FUNCTION "PDH_J_Raw" : Void
{ S7_Optimized_Access := 'TRUE' }
VERSION : 0.1
//Erzeugt vom PDH (PDH-Test) am 2026-11-15 10:00 UTC – bei Änderungen im PDH neu herunterladen.
//Datenbaustein "Daten", Variante mit Siemens-Bibliothek LMQTT (TLS möglich), S7-1500, höchstens 1024 Byte je Nachricht.
//Schreibt feste Zeichen (UTF-8) ab buf[pos]. Passt es nicht, wird ovf gesetzt und nichts geschrieben.
   VAR_INPUT
      s : String;
   END_VAR

   VAR_IN_OUT
      buf : Array[*] of Byte;
      pos : DInt;
      ovf : Bool;
   END_VAR

   VAR_TEMP
      i : Int;
      n : Int;
   END_VAR


BEGIN
	IF #ovf THEN
	    RETURN;
	END_IF;
	#n := LEN(#s);
	IF #pos < LOWER_BOUND(ARR := #buf, DIM := 1) OR #pos + INT_TO_DINT(#n) - 1 > UPPER_BOUND(ARR := #buf, DIM := 1) THEN
	    #ovf := TRUE;
	    RETURN;
	END_IF;
	FOR #i := 1 TO #n DO
	    #buf[#pos] := CHAR_TO_BYTE(#s[#i]);
	    #pos := #pos + 1;
	END_FOR;
END_FUNCTION

FUNCTION "PDH_J_DInt" : Void
{ S7_Optimized_Access := 'TRUE' }
VERSION : 0.1
//Erzeugt vom PDH (PDH-Test) am 2026-11-15 10:00 UTC – bei Änderungen im PDH neu herunterladen.
//Datenbaustein "Daten", Variante mit Siemens-Bibliothek LMQTT (TLS möglich), S7-1500, höchstens 1024 Byte je Nachricht.
//Schreibt v als Dezimalzahl (auch -2147483648).
   VAR_INPUT
      v : DInt;
   END_VAR

   VAR_IN_OUT
      buf : Array[*] of Byte;
      pos : DInt;
      ovf : Bool;
   END_VAR

   VAR_TEMP
      x : DInt;
      d : DInt;
      k : Int;
      i : Int;
      need : DInt;
      dig : Array[0..9] of Byte;
   END_VAR


BEGIN
	IF #ovf THEN
	    RETURN;
	END_IF;
	// Ziffern rückwärts sammeln, ohne das Vorzeichen umzudrehen (sonst Überlauf bei -2147483648)
	#x := #v;
	#k := 0;
	REPEAT
	    #d := #x MOD 10;
	    IF #d < 0 THEN
	        #d := -#d;
	    END_IF;
	    #dig[#k] := DINT_TO_BYTE(#d + 48);
	    #k := #k + 1;
	    #x := #x / 10;
	UNTIL #x = 0
	END_REPEAT;
	#need := INT_TO_DINT(#k);
	IF #v < 0 THEN
	    #need := #need + 1;
	END_IF;
	IF #pos < LOWER_BOUND(ARR := #buf, DIM := 1) OR #pos + #need - 1 > UPPER_BOUND(ARR := #buf, DIM := 1) THEN
	    #ovf := TRUE;
	    RETURN;
	END_IF;
	IF #v < 0 THEN
	    #buf[#pos] := 16#2D;   // -
	    #pos := #pos + 1;
	END_IF;
	FOR #i := #k - 1 TO 0 BY -1 DO
	    #buf[#pos] := #dig[#i];
	    #pos := #pos + 1;
	END_FOR;
END_FUNCTION

FUNCTION "PDH_J_UDInt" : Void
{ S7_Optimized_Access := 'TRUE' }
VERSION : 0.1
//Erzeugt vom PDH (PDH-Test) am 2026-11-15 10:00 UTC – bei Änderungen im PDH neu herunterladen.
//Datenbaustein "Daten", Variante mit Siemens-Bibliothek LMQTT (TLS möglich), S7-1500, höchstens 1024 Byte je Nachricht.
//Schreibt v als Dezimalzahl ohne Vorzeichen.
   VAR_INPUT
      v : UDInt;
   END_VAR

   VAR_IN_OUT
      buf : Array[*] of Byte;
      pos : DInt;
      ovf : Bool;
   END_VAR

   VAR_TEMP
      x : UDInt;
      k : Int;
      i : Int;
      dig : Array[0..9] of Byte;
   END_VAR


BEGIN
	IF #ovf THEN
	    RETURN;
	END_IF;
	#x := #v;
	#k := 0;
	REPEAT
	    #dig[#k] := UDINT_TO_BYTE(#x MOD 10 + 48);
	    #k := #k + 1;
	    #x := #x / 10;
	UNTIL #x = 0
	END_REPEAT;
	IF #pos < LOWER_BOUND(ARR := #buf, DIM := 1) OR #pos + INT_TO_DINT(#k) - 1 > UPPER_BOUND(ARR := #buf, DIM := 1) THEN
	    #ovf := TRUE;
	    RETURN;
	END_IF;
	FOR #i := #k - 1 TO 0 BY -1 DO
	    #buf[#pos] := #dig[#i];
	    #pos := #pos + 1;
	END_FOR;
END_FUNCTION

FUNCTION "PDH_J_Num" : Void
{ S7_Optimized_Access := 'TRUE' }
VERSION : 0.1
//Erzeugt vom PDH (PDH-Test) am 2026-11-15 10:00 UTC – bei Änderungen im PDH neu herunterladen.
//Datenbaustein "Daten", Variante mit Siemens-Bibliothek LMQTT (TLS möglich), S7-1500, höchstens 1024 Byte je Nachricht.
//Schreibt x mit digits gültigen Stellen wie Go strconv.FormatFloat(x, 'E', digits - 1, …):
//[-]d.ddd…E±XX, Exponent mit mindestens zwei Ziffern. NaN, ±unendlich und Beträge über maxAbs als null.
//Gerundet wird zur nächsten Zahl, bei genau der Mitte zur geraden. Für Beträge von 1E-8 bis 1E36
//wird der Rundungsfehler exakt mitgerechnet (Dekker); außerhalb kann die letzte Stelle selten abweichen.
//Gleich halten mit sclNum in generate_test.go (Go-Nachbau dieses Ablaufs).
   VAR_INPUT
      x : LReal;
      digits : Int;   // 7 für Real, 15 für LReal
      maxAbs : LReal;   // größter Betrag, der als Zahl geschrieben wird
   END_VAR

   VAR_IN_OUT
      buf : Array[*] of Byte;
      pos : DInt;
      ovf : Bool;
   END_VAR

   VAR_TEMP
      a : LReal;
      t : LReal;
      s : LReal;
      p : LReal;
      y : LReal;
      lo : LReal;
      n : LReal;
      f : LReal;
      top : LReal;
      c : LReal;
      ah : LReal;
      al : LReal;
      bh : LReal;
      bl : LReal;
      ph : LReal;
      e : Int;
      k : Int;
      j : Int;
      i : Int;
      pass : Int;
      hiD : DInt;
      loD : DInt;
      neg : Bool;
      exact : Bool;
      odd : Bool;
      dig : Array[1..15] of Byte;
   END_VAR


BEGIN
	IF #ovf THEN
	    RETURN;
	END_IF;
	IF #digits < 1 OR #digits > 15 OR #pos < LOWER_BOUND(ARR := #buf, DIM := 1) OR #pos + INT_TO_DINT(#digits) + 6 > UPPER_BOUND(ARR := #buf, DIM := 1) THEN
	    #ovf := TRUE;
	    RETURN;
	END_IF;
	// NaN, ±unendlich und zu große Beträge: null (jeder Vergleich mit NaN ist falsch)
	IF NOT (ABS(#x) <= #maxAbs) THEN
	    #buf[#pos] := 16#6E;   // n
	    #buf[#pos + 1] := 16#75;   // u
	    #buf[#pos + 2] := 16#6C;   // l
	    #buf[#pos + 3] := 16#6C;   // l
	    #pos := #pos + 4;
	    RETURN;
	END_IF;
	#neg := #x < 0.0;
	#a := ABS(#x);
	#top := 1.0;
	FOR #i := 1 TO #digits DO
	    #top := #top * 10.0;
	END_FOR;
	#n := 0.0;
	#e := 0;
	IF #a > 0.0 THEN
	    // Zehnerexponent schätzen (1 <= a / 10^e < 10), wird unten nachgebessert
	    #t := #a;
	    IF #t >= 1.0 THEN
	        IF #t >= LREAL#1.0E256 THEN #t := #t / LREAL#1.0E256; #e := #e + 256; END_IF;
	        IF #t >= LREAL#1.0E128 THEN #t := #t / LREAL#1.0E128; #e := #e + 128; END_IF;
	        IF #t >= LREAL#1.0E64 THEN #t := #t / LREAL#1.0E64; #e := #e + 64; END_IF;
	        IF #t >= LREAL#1.0E32 THEN #t := #t / LREAL#1.0E32; #e := #e + 32; END_IF;
	        IF #t >= LREAL#1.0E16 THEN #t := #t / LREAL#1.0E16; #e := #e + 16; END_IF;
	        IF #t >= LREAL#1.0E8 THEN #t := #t / LREAL#1.0E8; #e := #e + 8; END_IF;
	        IF #t >= LREAL#1.0E4 THEN #t := #t / LREAL#1.0E4; #e := #e + 4; END_IF;
	        IF #t >= LREAL#1.0E2 THEN #t := #t / LREAL#1.0E2; #e := #e + 2; END_IF;
	        IF #t >= LREAL#1.0E1 THEN #t := #t / LREAL#1.0E1; #e := #e + 1; END_IF;
	    ELSE
	        IF #t < LREAL#1.0E-255 THEN #t := #t * LREAL#1.0E256; #e := #e - 256; END_IF;
	        IF #t < LREAL#1.0E-127 THEN #t := #t * LREAL#1.0E128; #e := #e - 128; END_IF;
	        IF #t < LREAL#1.0E-63 THEN #t := #t * LREAL#1.0E64; #e := #e - 64; END_IF;
	        IF #t < LREAL#1.0E-31 THEN #t := #t * LREAL#1.0E32; #e := #e - 32; END_IF;
	        IF #t < LREAL#1.0E-15 THEN #t := #t * LREAL#1.0E16; #e := #e - 16; END_IF;
	        IF #t < LREAL#1.0E-7 THEN #t := #t * LREAL#1.0E8; #e := #e - 8; END_IF;
	        IF #t < LREAL#1.0E-3 THEN #t := #t * LREAL#1.0E4; #e := #e - 4; END_IF;
	        IF #t < LREAL#1.0E-1 THEN #t := #t * LREAL#1.0E2; #e := #e - 2; END_IF;
	        IF #t < LREAL#1.0 THEN #t := #t * LREAL#1.0E1; #e := #e - 1; END_IF;
	    END_IF;
	    // Mantisse n = a * 10^k als ganze Zahl mit digits Stellen
	    FOR #pass := 1 TO 3 DO
	        #k := #digits - 1 - #e;
	        IF #k > 300 THEN
	            // sehr kleine Zahlen: 10^k läge über dem LReal-Bereich
	            #s := #a * LREAL#1.0E100;
	            #j := #k - 100;
	        ELSE
	            #s := #a;
	            #j := ABS(#k);
	        END_IF;
	        #p := 1.0;
	        IF #j >= 256 THEN #p := #p * LREAL#1.0E256; #j := #j - 256; END_IF;
	        IF #j >= 128 THEN #p := #p * LREAL#1.0E128; #j := #j - 128; END_IF;
	        IF #j >= 64 THEN #p := #p * LREAL#1.0E64; #j := #j - 64; END_IF;
	        IF #j >= 32 THEN #p := #p * LREAL#1.0E32; #j := #j - 32; END_IF;
	        IF #j >= 16 THEN #p := #p * LREAL#1.0E16; #j := #j - 16; END_IF;
	        IF #j >= 8 THEN #p := #p * LREAL#1.0E8; #j := #j - 8; END_IF;
	        IF #j >= 4 THEN #p := #p * LREAL#1.0E4; #j := #j - 4; END_IF;
	        IF #j >= 2 THEN #p := #p * LREAL#1.0E2; #j := #j - 2; END_IF;
	        IF #j >= 1 THEN #p := #p * LREAL#1.0E1; #j := #j - 1; END_IF;
	        // bis 10^22 ist p exakt, dann lässt sich der Rundungsfehler lo exakt bestimmen
	        #exact := #k >= -22 AND #k <= 22;
	        #lo := 0.0;
	        IF #k >= 0 THEN
	            #y := #s * #p;
	            IF #exact THEN
	                // Fehler der Multiplikation (Dekker, Teilung mit 2^27 + 1)
	                #c := LREAL#134217729.0 * #s;
	                #ah := #c - (#c - #s);
	                #al := #s - #ah;
	                #c := LREAL#134217729.0 * #p;
	                #bh := #c - (#c - #p);
	                #bl := #p - #bh;
	                #lo := (((#ah * #bh - #y) + #ah * #bl) + #al * #bh) + #al * #bl;
	            END_IF;
	        ELSE
	            #y := #s / #p;
	            IF #exact THEN
	                // Rest der Division s - y * p exakt, dann durch p
	                #ph := #y * #p;
	                #c := LREAL#134217729.0 * #y;
	                #ah := #c - (#c - #y);
	                #al := #y - #ah;
	                #c := LREAL#134217729.0 * #p;
	                #bh := #c - (#c - #p);
	                #bl := #p - #bh;
	                #lo := (((#ah * #bh - #ph) + #ah * #bl) + #al * #bh) + #al * #bl;
	                #lo := ((#s - #ph) - #lo) / #p;
	            END_IF;
	        END_IF;
	        // zur nächsten ganzen Zahl runden: (y + 2^52) - 2^52, bei genau .5 zur geraden
	        #t := #y + LREAL#4503599627370496.0;
	        #n := #t - LREAL#4503599627370496.0;
	        #f := #y - #n;
	        #t := #n / 2.0 + LREAL#4503599627370496.0;
	        #odd := (#t - LREAL#4503599627370496.0) <> #n / 2.0;
	        IF #f = 0.5 AND (#lo > 0.0 OR (#lo = 0.0 AND #odd)) THEN
	            #n := #n + 1.0;
	        ELSIF #f = -0.5 AND (#lo < 0.0 OR (#lo = 0.0 AND #odd)) THEN
	            #n := #n - 1.0;
	        END_IF;
	        IF #n >= #top THEN
	            #e := #e + 1;
	        ELSIF #n < #top / 10.0 THEN
	            #e := #e - 1;
	        ELSE
	            EXIT;
	        END_IF;
	    END_FOR;
	    // über der größten LReal-Zahl, die PDH noch liest: null
	    IF #e = 308 AND #n > LREAL#179769313486231.0 THEN
	        #buf[#pos] := 16#6E;   // n
	        #buf[#pos + 1] := 16#75;   // u
	        #buf[#pos + 2] := 16#6C;   // l
	        #buf[#pos + 3] := 16#6C;   // l
	        #pos := #pos + 4;
	        RETURN;
	    END_IF;
	END_IF;
	// Ziffern: n = hiD * 10^8 + loD
	#hiD := TRUNC(#n / LREAL#1.0E8);
	#loD := LREAL_TO_DINT(#n - DINT_TO_LREAL(#hiD) * LREAL#1.0E8);
	IF #loD < 0 THEN
	    #hiD := #hiD - 1;
	    #loD := #loD + 100000000;
	ELSIF #loD >= 100000000 THEN
	    #hiD := #hiD + 1;
	    #loD := #loD - 100000000;
	END_IF;
	FOR #i := #digits TO 1 BY -1 DO
	    IF #digits - #i < 8 THEN
	        #dig[#i] := DINT_TO_BYTE(#loD MOD 10 + 48);
	        #loD := #loD / 10;
	    ELSE
	        #dig[#i] := DINT_TO_BYTE(#hiD MOD 10 + 48);
	        #hiD := #hiD / 10;
	    END_IF;
	END_FOR;
	IF #neg THEN
	    #buf[#pos] := 16#2D;   // -
	    #pos := #pos + 1;
	END_IF;
	#buf[#pos] := #dig[1];
	#buf[#pos + 1] := 16#2E;   // .
	#pos := #pos + 2;
	FOR #i := 2 TO #digits DO
	    #buf[#pos] := #dig[#i];
	    #pos := #pos + 1;
	END_FOR;
	#buf[#pos] := 16#45;   // E
	IF #e < 0 THEN
	    #buf[#pos + 1] := 16#2D;   // -
	    #e := -#e;
	ELSE
	    #buf[#pos + 1] := 16#2B;   // +
	END_IF;
	#pos := #pos + 2;
	IF #e >= 100 THEN
	    #buf[#pos] := INT_TO_BYTE(#e / 100 + 48);
	    #pos := #pos + 1;
	END_IF;
	#buf[#pos] := INT_TO_BYTE((#e / 10) MOD 10 + 48);
	#buf[#pos + 1] := INT_TO_BYTE(#e MOD 10 + 48);
	#pos := #pos + 2;
END_FUNCTION

FUNCTION "PDH_J_Real" : Void
{ S7_Optimized_Access := 'TRUE' }
VERSION : 0.1
//Erzeugt vom PDH (PDH-Test) am 2026-11-15 10:00 UTC – bei Änderungen im PDH neu herunterladen.
//Datenbaustein "Daten", Variante mit Siemens-Bibliothek LMQTT (TLS möglich), S7-1500, höchstens 1024 Byte je Nachricht.
//Schreibt v wie Go strconv.FormatFloat(v, 'E', 6, 32), z. B. 1.450000E+03; NaN und ±unendlich als null.
   VAR_INPUT
      v : Real;
   END_VAR

   VAR_IN_OUT
      buf : Array[*] of Byte;
      pos : DInt;
      ovf : Bool;
   END_VAR


BEGIN
	"PDH_J_Num"(x := REAL_TO_LREAL(#v), digits := 7, maxAbs := LREAL#3.4028234663852886E+38, buf := #buf, pos := #pos, ovf := #ovf);
END_FUNCTION

FUNCTION "PDH_J_LReal" : Void
{ S7_Optimized_Access := 'TRUE' }
VERSION : 0.1
//Erzeugt vom PDH (PDH-Test) am 2026-11-15 10:00 UTC – bei Änderungen im PDH neu herunterladen.
//Datenbaustein "Daten", Variante mit Siemens-Bibliothek LMQTT (TLS möglich), S7-1500, höchstens 1024 Byte je Nachricht.
//Schreibt v wie Go strconv.FormatFloat(v, 'E', 14, 64); NaN, ±unendlich und Beträge über 1.79769313486231E+308 als null.
   VAR_INPUT
      v : LReal;
   END_VAR

   VAR_IN_OUT
      buf : Array[*] of Byte;
      pos : DInt;
      ovf : Bool;
   END_VAR


BEGIN
	"PDH_J_Num"(x := #v, digits := 15, maxAbs := LREAL#1.79769313486231E+308, buf := #buf, pos := #pos, ovf := #ovf);
END_FUNCTION

FUNCTION "PDH_J_Str" : Void
{ S7_Optimized_Access := 'TRUE' }
VERSION : 0.1
//Erzeugt vom PDH (PDH-Test) am 2026-11-15 10:00 UTC – bei Änderungen im PDH neu herunterladen.
//Datenbaustein "Daten", Variante mit Siemens-Bibliothek LMQTT (TLS möglich), S7-1500, höchstens 1024 Byte je Nachricht.
//Schreibt s als JSON-Zeichenkette: " und \ mit \ davor, Steuerzeichen als Leerzeichen,
//Zeichen ab 16#80 (Latin-1) als zwei Byte UTF-8.
   VAR_INPUT
      s : String;
   END_VAR

   VAR_IN_OUT
      buf : Array[*] of Byte;
      pos : DInt;
      ovf : Bool;
   END_VAR

   VAR_TEMP
      i : Int;
      n : Int;
      b : Byte;
      c : Int;
   END_VAR


BEGIN
	IF #ovf THEN
	    RETURN;
	END_IF;
	#n := LEN(#s);
	// je Zeichen höchstens zwei Byte, dazu die Anführungszeichen
	IF #pos < LOWER_BOUND(ARR := #buf, DIM := 1) OR #pos + 2 * INT_TO_DINT(#n) + 1 > UPPER_BOUND(ARR := #buf, DIM := 1) THEN
	    #ovf := TRUE;
	    RETURN;
	END_IF;
	#buf[#pos] := 16#22;   // "
	#pos := #pos + 1;
	FOR #i := 1 TO #n DO
	    #b := CHAR_TO_BYTE(#s[#i]);
	    #c := BYTE_TO_INT(#b);
	    IF #c = 34 OR #c = 92 THEN
	        #buf[#pos] := 16#5C;   // \
	        #buf[#pos + 1] := #b;
	        #pos := #pos + 2;
	    ELSIF #c < 32 THEN
	        #buf[#pos] := 16#20;
	        #pos := #pos + 1;
	    ELSIF #c < 128 THEN
	        #buf[#pos] := #b;
	        #pos := #pos + 1;
	    ELSE
	        #buf[#pos] := INT_TO_BYTE(192 + #c / 64);
	        #buf[#pos + 1] := INT_TO_BYTE(128 + #c MOD 64);
	        #pos := #pos + 2;
	    END_IF;
	END_FOR;
	#buf[#pos] := 16#22;   // "
	#pos := #pos + 1;
END_FUNCTION

FUNCTION "PDH_J_DTL" : Void
{ S7_Optimized_Access := 'TRUE' }
VERSION : 0.1
//Erzeugt vom PDH (PDH-Test) am 2026-11-15 10:00 UTC – bei Änderungen im PDH neu herunterladen.
//Datenbaustein "Daten", Variante mit Siemens-Bibliothek LMQTT (TLS möglich), S7-1500, höchstens 1024 Byte je Nachricht.
//Schreibt v als "JJJJ-MM-TTThh:mm:ss", mit zone = TRUE als "JJJJ-MM-TTThh:mm:ssZ" (UTC).
   VAR_INPUT
      v : DTL;
      zone : Bool;
   END_VAR

   VAR_IN_OUT
      buf : Array[*] of Byte;
      pos : DInt;
      ovf : Bool;
   END_VAR

   VAR_TEMP
      f : Int;
      i : Int;
      w : Int;
      x : DInt;
      sep : Byte;
   END_VAR


BEGIN
	IF #ovf THEN
	    RETURN;
	END_IF;
	IF #pos < LOWER_BOUND(ARR := #buf, DIM := 1) OR #pos + 21 > UPPER_BOUND(ARR := #buf, DIM := 1) THEN
	    #ovf := TRUE;
	    RETURN;
	END_IF;
	#buf[#pos] := 16#22;   // "
	#pos := #pos + 1;
	FOR #f := 1 TO 6 DO
	    CASE #f OF
	        1:
	            #x := UINT_TO_DINT(#v.YEAR);
	            #w := 4;
	            #sep := 16#2D;   // -
	        2:
	            #x := USINT_TO_DINT(#v.MONTH);
	            #w := 2;
	            #sep := 16#2D;   // -
	        3:
	            #x := USINT_TO_DINT(#v.DAY);
	            #w := 2;
	            #sep := 16#54;   // T
	        4:
	            #x := USINT_TO_DINT(#v.HOUR);
	            #w := 2;
	            #sep := 16#3A;   // :
	        5:
	            #x := USINT_TO_DINT(#v.MINUTE);
	            #w := 2;
	            #sep := 16#3A;   // :
	        ELSE
	            #x := USINT_TO_DINT(#v.SECOND);
	            #w := 2;
	            #sep := 16#22;   // "
	    END_CASE;
	    FOR #i := #w - 1 TO 0 BY -1 DO
	        #buf[#pos + #i] := DINT_TO_BYTE(#x MOD 10 + 48);
	        #x := #x / 10;
	    END_FOR;
	    #pos := #pos + #w;
	    IF #f < 6 THEN
	        #buf[#pos] := #sep;
	        #pos := #pos + 1;
	    END_IF;
	END_FOR;
	IF #zone THEN
	    #buf[#pos] := 16#5A;   // Z
	    #pos := #pos + 1;
	END_IF;
	#buf[#pos] := 16#22;   // "
	#pos := #pos + 1;
END_FUNCTION

FUNCTION_BLOCK "PDH_MQTT_Daten"
{ S7_Optimized_Access := 'TRUE' }
VERSION : 0.1
//Erzeugt vom PDH (PDH-Test) am 2026-11-15 10:00 UTC – bei Änderungen im PDH neu herunterladen.
//Datenbaustein "Daten", Variante mit Siemens-Bibliothek LMQTT (TLS möglich), S7-1500, höchstens 1024 Byte je Nachricht.
//Sendet die Werte aus "daten" per MQTT (QoS 0) an den Broker aus "PDH_Daten_Konfig":
//bei steigender Flanke an trigger als 2 Nachricht(en), dazu regelmäßig einen Heartbeat.
//Nutzt den FB "LMQTT_Client" der Siemens-Bibliothek LMQTT (TLS möglich). Je Verbindung nur einmal aufrufen.
//
//Vor dem Einsatz mit der Doku der eingesetzten LMQTT-Version abgleichen (erstellt nach
//Beitrag 109748872 V3.1 04/2024, "LMQTT_Client" V4.0.4):
//  Baustein "LMQTT_Client", Datentyp "LMQTT_typeConnParam" mit hwId, connId, broker, port,
//  tls.enableTls, tls.validateServerIdentity, tls.brokerCert, tls.clientCert, keepAlive;
//  Parameter enable, publish, subscribe, unsubscribe, connParam, clientIdentifier, username,
//  password, willTopic, willMsgPayload, willMsgLen, qos, mqttTopic, publishMsgPayload,
//  publishMsgLen, retain, receivedTopic, receivedMsgPayload, receivedMsgDataLen,
//  receivedMsgStatus; Ausgänge done, error, status; Bibliotheksstatus (instClient.status)
//  16#7003 TCP verbunden, 16#7004 MQTT verbunden, 16#9000 Verbindung unterbrochen.
   VAR_INPUT
      enable : Bool;   // TRUE = verbinden und bereit halten
      trigger : Bool;   // steigende Flanke = Werte senden
      heartbeatInterval : Time := T#60s;   // T#0s = kein Heartbeat
      hwId : HW_ANY := 64;   // Hardware-Kennung der PROFINET-Schnittstelle
      connId : CONN_OUC := 1;   // Verbindungsnummer, in der Steuerung eindeutig
   END_VAR

   VAR_OUTPUT
      connected : Bool;
      busy : Bool;
      done : Bool;   // einen Zyklus nach dem letzten Teil
      error : Bool;
      status : Word;
      statusText : String[60];
      sentCount : UDInt;
      heartbeatCount : UDInt;
   END_VAR

   VAR_IN_OUT
      daten : "PDH_Daten_Typ";
   END_VAR

   VAR
      snap : "PDH_Daten_Typ";   // Abbild der Werte beim Trigger
      ts : DTL;   // Zeitstempel (UTC) aller Teile eines Triggers
      hbTs : DTL;
      pl : Array[0..1023] of Byte;   // JSON-Inhalt einer Nachricht
      instClient : "LMQTT_Client";   // Bibliothek LMQTT
      connParam : "LMQTT_typeConnParam";
      clientId : WString[254];
      user : WString[254];
      pass : WString[254];
      willTopic : WString[254];   // kein Last Will
      willMsg : Array[0..0] of Byte;
      willLen : UInt;
      qos : USInt;
      pubTopic : WString[254];
      pubLen : UDInt;
      pubRetain : Bool;
      rxTopic : WString[200];   // Empfang wird nicht genutzt
      rxMsg : Array[0..0] of Byte;
      rxLen : UDInt;
      rxStatus : USInt;
      trigEdge : R_TRIG;
      tmrConn : TON;
      tmrSend : TON;
      tmrRetry : TON;
      tmrHb : TON;
      state : Int;
      buildKind : Int;
      sendKind : Int;
      part : Int;
      pos : DInt;
      ovf : Bool;
      libEnable : Bool;
      libUp : Bool;
      libStatus : Word;
      pubReq : Bool;
      failed : Bool;
      failCode : Word;
      failText : String[60];
      lastErr : Word;
      lastText : String[60];
      evStatus : Word;
      evText : String[60];
      trigPending : Bool;
      hbDue : Bool;
   END_VAR

   VAR_TEMP
      i : Int;
      n : Int;
      c : Int;
      rc : Int;
   END_VAR


BEGIN
	// ---------------------------------------------------------------- Zyklusanfang
	#done := FALSE;
	#error := FALSE;
	#evStatus := 16#0000;
	#failCode := 16#0000;
	#buildKind := 0;

	// Zeitglieder jeden Zyklus aufrufen, dann laufen sie beim Zustandswechsel neu an.
	#tmrConn(IN := (#state = 1), PT := T#30s);
	#tmrSend(IN := (#state = 4 AND #pubReq), PT := T#10s);
	#tmrRetry(IN := (#state = 6), PT := T#5s);
	#tmrHb(IN := (#connected AND #heartbeatInterval > T#0s AND NOT #hbDue), PT := #heartbeatInterval);
	IF #tmrHb.Q THEN
	    #hbDue := TRUE;
	END_IF;

	// ---------------------------------------------------------------- Trigger
	#trigEdge(CLK := #trigger);
	IF #trigEdge.Q THEN
	    IF #connected AND #enable THEN
	        // wird in "bereit" gestartet; während busy bleibt genau eine Wiederholung gemerkt
	        #trigPending := TRUE;
	    ELSE
	        // nicht verbunden: nichts puffern
	        #evStatus := 16#8007;
	        #evText := 'nicht verbunden beim Trigger';
	    END_IF;
	END_IF;

	// ---------------------------------------------------------------- Bibliothek LMQTT
	IF #state = 1 AND NOT #libEnable THEN
	    // Verbindungsdaten beim (Neu-)Verbinden aus der Konfiguration übernehmen
	    #connParam.hwId := #hwId;
	    #connParam.connId := #connId;
	    #connParam.broker := "PDH_Daten_Konfig".brokerHost;
	    #connParam.port := "PDH_Daten_Konfig".brokerPort;
	    #connParam.tls.enableTls := "PDH_Daten_Konfig".useTls;
	    #connParam.tls.validateServerIdentity := "PDH_Daten_Konfig".validateServer;
	    #connParam.tls.brokerCert := "PDH_Daten_Konfig".brokerCert;
	    #connParam.tls.clientCert := "PDH_Daten_Konfig".clientCert;
	    #connParam.keepAlive := "PDH_Daten_Konfig".keepAlive;
	    #clientId := "PDH_Daten_Konfig".clientId;
	    #user := "PDH_Daten_Konfig".username;
	    #pass := "PDH_Daten_Konfig".password;
	    #willTopic := WSTRING#'';
	    #willLen := 0;
	    #qos := 0;   // QoS 0 wie die eigenständige Variante
	    #libEnable := TRUE;   // steigende Flanke an enable: Bibliothek verbindet
	END_IF;
	#instClient(enable := #libEnable,
	            publish := #pubReq,
	            subscribe := FALSE,
	            unsubscribe := FALSE,
	            connParam := #connParam,
	            clientIdentifier := #clientId,
	            username := #user,
	            password := #pass,
	            willTopic := #willTopic,
	            willMsgPayload := #willMsg,
	            willMsgLen := #willLen,
	            qos := #qos,
	            mqttTopic := #pubTopic,
	            publishMsgPayload := #pl,
	            publishMsgLen := #pubLen,
	            retain := #pubRetain,
	            receivedTopic := #rxTopic,
	            receivedMsgPayload := #rxMsg,
	            receivedMsgDataLen := #rxLen,
	            receivedMsgStatus := #rxStatus);
	#libStatus := #instClient.status;
	IF NOT #libEnable THEN
	    #libUp := FALSE;
	ELSIF #instClient.error THEN
	    // Fehler der Bibliothek: 16#82xx, ihr Status steht als 16#xxxx am Ende von statusText
	    IF #state = 4 THEN
	        #failCode := 16#8202;
	        #failText := 'LMQTT Sendefehler 16#0000';
	    ELSE
	        #failCode := 16#8201;
	        #failText := 'LMQTT Verbindungsfehler 16#0000';
	    END_IF;
	    #n := LEN(#failText) - 4;
	    FOR #i := 1 TO 4 DO
	        #c := WORD_TO_INT(SHR(IN := #libStatus, N := 16 - 4 * #i) AND 16#000F);
	        IF #c < 10 THEN
	            #c := #c + 48;
	        ELSE
	            #c := #c + 55;
	        END_IF;
	        #failText[#n + #i] := BYTE_TO_CHAR(INT_TO_BYTE(#c));
	    END_FOR;
	ELSIF #libStatus = 16#7004 THEN
	    #libUp := TRUE;   // MQTT verbunden, kein Auftrag aktiv
	ELSIF #libStatus = 16#9000 OR #libStatus = 16#7000 OR #libStatus = 16#7001 OR #libStatus = 16#7002 OR #libStatus = 16#7003 THEN
	    #libUp := FALSE;   // unterbrochen oder noch nicht angemeldet
	END_IF;

	// ---------------------------------------------------------------- Verbindung unterbrochen
	// Die Bibliothek verbindet selbst neu. Wie bei einem Fehler wird nichts Gemerktes
	// (Trigger, Heartbeat) über die Unterbrechung mitgenommen.
	IF (#state = 3 OR #state = 4) AND NOT #libUp AND #failCode = 16#0000 THEN
	    IF #state = 4 THEN
	        #evStatus := 16#8002;
	        #evText := 'Sendefehler (Verbindung unterbrochen)';
	    END_IF;
	    #connected := FALSE;
	    #busy := FALSE;
	    #trigPending := FALSE;
	    #hbDue := FALSE;
	    #pubReq := FALSE;
	    #state := 1;
	END_IF;

	// ---------------------------------------------------------------- Ablauf
	IF #failCode = 16#0000 THEN
	    CASE #state OF
	        0:  // aus
	            #connected := FALSE;
	            #busy := FALSE;
	            #failed := FALSE;
	            #libEnable := FALSE;
	            #pubReq := FALSE;
	            #trigPending := FALSE;
	            #hbDue := FALSE;
	            IF #enable THEN
	                #state := 1;
	            END_IF;

	        1:  // verbinden (TCP/TLS und MQTT macht die Bibliothek)
	            IF NOT #enable THEN
	                #libEnable := FALSE;
	                #state := 6;
	            ELSIF #libUp THEN
	                #connected := TRUE;
	                #failed := FALSE;
	                #state := 3;
	            ELSIF #tmrConn.Q THEN
	                #failCode := 16#8005;
	                #failText := 'keine Antwort vom Broker';
	            END_IF;

	        3:  // bereit
	            IF NOT #enable THEN
	                #libEnable := FALSE;
	                #connected := FALSE;
	                #state := 6;
	            ELSIF #trigPending THEN
	                #trigPending := FALSE;
	                #rc := RD_SYS_T(OUT => #ts);
	                IF #rc <> 0 THEN
	                    #evStatus := 16#8009;
	                    #evText := 'Uhrzeit nicht lesbar';
	                ELSE
	                    #snap := #daten;   // alle Teile aus demselben Abbild
	                    #part := 1;
	                    #busy := TRUE;
	                    #buildKind := 2;
	                END_IF;
	            ELSIF #hbDue THEN
	                #rc := RD_SYS_T(OUT => #hbTs);
	                IF #rc <> 0 THEN
	                    #hbDue := FALSE;
	                    #evStatus := 16#8009;
	                    #evText := 'Uhrzeit nicht lesbar';
	                ELSE
	                    #buildKind := 3;
	                END_IF;
	            END_IF;

	        4:  // senden: publish bleibt TRUE bis done, dann mindestens einen Zyklus FALSE
	            IF NOT #pubReq THEN
	                // publish war einen Zyklus FALSE: nächsten Teil bauen
	                #buildKind := 2;
	            ELSIF #instClient.done THEN
	                #pubReq := FALSE;   // zurücknehmen, sonst bleibt done stehen
	                CASE #sendKind OF
	                    2:  // Teil
	                        IF #part < 2 AND #enable THEN
	                            #part := #part + 1;   // im nächsten Zyklus bauen, publish ist dann einen Zyklus FALSE
	                        ELSE
	                            IF #part >= 2 THEN
	                                #done := TRUE;
	                                #sentCount := #sentCount + 1;
	                            END_IF;
	                            #busy := FALSE;
	                            #state := 3;
	                        END_IF;
	                    3:  // Heartbeat
	                        #heartbeatCount := #heartbeatCount + 1;
	                        #hbDue := FALSE;
	                        #state := 3;
	                END_CASE;
	            ELSIF #tmrSend.Q THEN
	                #failCode := 16#8002;
	                #failText := 'Sendefehler (keine Antwort)';
	            END_IF;

	        6:  // Bibliothek aus, 5 s warten, dann neu verbinden
	            #connected := FALSE;
	            #busy := FALSE;
	            #libEnable := FALSE;
	            #pubReq := FALSE;
	            IF #tmrRetry.Q THEN
	                IF #enable THEN
	                    #state := 1;
	                ELSE
	                    #state := 0;
	                END_IF;
	            END_IF;

	        ELSE
	            #state := 0;
	    END_CASE;
	END_IF;

	// ---------------------------------------------------------------- Nachricht bauen
	IF #buildKind <> 0 AND #failCode = 16#0000 THEN
	    #ovf := FALSE;
	    #pos := 0;
	    CASE #buildKind OF
	        2:  // Teil #part: JSON in #pl
	            "PDH_J_Raw"(s := '{"ts":', buf := #pl, pos := #pos, ovf := #ovf);
	            "PDH_J_DTL"(v := #ts, zone := TRUE, buf := #pl, pos := #pos, ovf := #ovf);
	            "PDH_J_Raw"(s := ',"part":', buf := #pl, pos := #pos, ovf := #ovf);
	            "PDH_J_DInt"(v := INT_TO_DINT(#part), buf := #pl, pos := #pos, ovf := #ovf);
	            "PDH_J_Raw"(s := ',"parts":2,"values":{', buf := #pl, pos := #pos, ovf := #ovf);
	            CASE #part OF
	                1:
	                    "PDH_J_Raw"(s := '"Zaehler":', buf := #pl, pos := #pos, ovf := #ovf);
	                    "PDH_J_Real"(v := #snap."Zaehler", buf := #pl, pos := #pos, ovf := #ovf);
	                    "PDH_J_Raw"(s := ',"Takt":', buf := #pl, pos := #pos, ovf := #ovf);
	                    "PDH_J_DInt"(v := INT_TO_DINT(#snap."Takt"), buf := #pl, pos := #pos, ovf := #ovf);
	                    "PDH_J_Raw"(s := ',"Motor":{"Drehzahl":', buf := #pl, pos := #pos, ovf := #ovf);
	                    "PDH_J_Real"(v := #snap."Motor"."Drehzahl", buf := #pl, pos := #pos, ovf := #ovf);
	                    "PDH_J_Raw"(s := ',"Ein":', buf := #pl, pos := #pos, ovf := #ovf);
	                    IF #snap."Motor"."Ein" THEN
	                        "PDH_J_Raw"(s := 'true', buf := #pl, pos := #pos, ovf := #ovf);
	                    ELSE
	                        "PDH_J_Raw"(s := 'false', buf := #pl, pos := #pos, ovf := #ovf);
	                    END_IF;
	                    "PDH_J_Raw"(s := '},"Feld":[', buf := #pl, pos := #pos, ovf := #ovf);
	                    "PDH_J_DInt"(v := INT_TO_DINT(#snap."Feld"[1]), buf := #pl, pos := #pos, ovf := #ovf);
	                    "PDH_J_Raw"(s := ',', buf := #pl, pos := #pos, ovf := #ovf);
	                    "PDH_J_DInt"(v := INT_TO_DINT(#snap."Feld"[2]), buf := #pl, pos := #pos, ovf := #ovf);
	                    "PDH_J_Raw"(s := ',', buf := #pl, pos := #pos, ovf := #ovf);
	                    "PDH_J_DInt"(v := INT_TO_DINT(#snap."Feld"[3]), buf := #pl, pos := #pos, ovf := #ovf);
	                    "PDH_J_Raw"(s := ',', buf := #pl, pos := #pos, ovf := #ovf);
	                    "PDH_J_DInt"(v := INT_TO_DINT(#snap."Feld"[4]), buf := #pl, pos := #pos, ovf := #ovf);
	                    "PDH_J_Raw"(s := ',', buf := #pl, pos := #pos, ovf := #ovf);
	                    "PDH_J_DInt"(v := INT_TO_DINT(#snap."Feld"[5]), buf := #pl, pos := #pos, ovf := #ovf);
	                    "PDH_J_Raw"(s := ',', buf := #pl, pos := #pos, ovf := #ovf);
	                    "PDH_J_DInt"(v := INT_TO_DINT(#snap."Feld"[6]), buf := #pl, pos := #pos, ovf := #ovf);
	                    "PDH_J_Raw"(s := ',', buf := #pl, pos := #pos, ovf := #ovf);
	                    "PDH_J_DInt"(v := INT_TO_DINT(#snap."Feld"[7]), buf := #pl, pos := #pos, ovf := #ovf);
	                    "PDH_J_Raw"(s := ',', buf := #pl, pos := #pos, ovf := #ovf);
	                    "PDH_J_DInt"(v := INT_TO_DINT(#snap."Feld"[8]), buf := #pl, pos := #pos, ovf := #ovf);
	                    "PDH_J_Raw"(s := ',', buf := #pl, pos := #pos, ovf := #ovf);
	                    "PDH_J_DInt"(v := INT_TO_DINT(#snap."Feld"[9]), buf := #pl, pos := #pos, ovf := #ovf);
	                    "PDH_J_Raw"(s := ',', buf := #pl, pos := #pos, ovf := #ovf);
	                    "PDH_J_DInt"(v := INT_TO_DINT(#snap."Feld"[10]), buf := #pl, pos := #pos, ovf := #ovf);
	                    "PDH_J_Raw"(s := '],"Text":', buf := #pl, pos := #pos, ovf := #ovf);
	                    "PDH_J_Str"(s := #snap."Text", buf := #pl, pos := #pos, ovf := #ovf);
	                    "PDH_J_Raw"(s := ',"Name":', buf := #pl, pos := #pos, ovf := #ovf);
	                    "PDH_J_Str"(s := #snap."Name", buf := #pl, pos := #pos, ovf := #ovf);
	                    "PDH_J_Raw"(s := ',"Zeit":', buf := #pl, pos := #pos, ovf := #ovf);
	                    "PDH_J_DTL"(v := #snap."Zeit", zone := FALSE, buf := #pl, pos := #pos, ovf := #ovf);
	                    "PDH_J_Raw"(s := ',"Wort":', buf := #pl, pos := #pos, ovf := #ovf);
	                    "PDH_J_UDInt"(v := WORD_TO_UDINT(#snap."Wort"), buf := #pl, pos := #pos, ovf := #ovf);
	                    "PDH_J_Raw"(s := ',"Doppelwort":', buf := #pl, pos := #pos, ovf := #ovf);
	                    "PDH_J_UDInt"(v := DWORD_TO_UDINT(#snap."Doppelwort"), buf := #pl, pos := #pos, ovf := #ovf);
	                    "PDH_J_Raw"(s := ',"Ganz":', buf := #pl, pos := #pos, ovf := #ovf);
	                    "PDH_J_DInt"(v := #snap."Ganz", buf := #pl, pos := #pos, ovf := #ovf);
	                    "PDH_J_Raw"(s := ',"Vorzeichenlos":', buf := #pl, pos := #pos, ovf := #ovf);
	                    "PDH_J_UDInt"(v := UINT_TO_UDINT(#snap."Vorzeichenlos"), buf := #pl, pos := #pos, ovf := #ovf);
	                    "PDH_J_Raw"(s := ',"Gross":', buf := #pl, pos := #pos, ovf := #ovf);
	                    "PDH_J_UDInt"(v := #snap."Gross", buf := #pl, pos := #pos, ovf := #ovf);
	                    "PDH_J_Raw"(s := ',"Genau":', buf := #pl, pos := #pos, ovf := #ovf);
	                    "PDH_J_LReal"(v := #snap."Genau", buf := #pl, pos := #pos, ovf := #ovf);
	                    "PDH_J_Raw"(s := ',"Zeitstempel":', buf := #pl, pos := #pos, ovf := #ovf);
	                    "PDH_J_DTL"(v := DT_TO_DTL(#snap."Zeitstempel"), zone := FALSE, buf := #pl, pos := #pos, ovf := #ovf);
	                2:
	                    "PDH_J_Raw"(s := '"Bemerkung":', buf := #pl, pos := #pos, ovf := #ovf);
	                    "PDH_J_Str"(s := #snap."Bemerkung", buf := #pl, pos := #pos, ovf := #ovf);
	                    "PDH_J_Raw"(s := ',"Z$C3$A4hler":{"St$C3$BCck":', buf := #pl, pos := #pos, ovf := #ovf);
	                    "PDH_J_UDInt"(v := #snap."Zähler"."Stück", buf := #pl, pos := #pos, ovf := #ovf);
	                    "PDH_J_Raw"(s := ',"it$'s":', buf := #pl, pos := #pos, ovf := #ovf);
	                    IF #snap."Zähler"."it's" THEN
	                        "PDH_J_Raw"(s := 'true', buf := #pl, pos := #pos, ovf := #ovf);
	                    ELSE
	                        "PDH_J_Raw"(s := 'false', buf := #pl, pos := #pos, ovf := #ovf);
	                    END_IF;
	                    "PDH_J_Raw"(s := '}', buf := #pl, pos := #pos, ovf := #ovf);
	            END_CASE;
	            "PDH_J_Raw"(s := '}}', buf := #pl, pos := #pos, ovf := #ovf);
	            #pubTopic := "PDH_Daten_Konfig".topic;
	            #pubRetain := "PDH_Daten_Konfig".retain;   // Retain nur für die Werte

	        3:  // --- Heartbeat ---
	            "PDH_J_Raw"(s := '{"ts":', buf := #pl, pos := #pos, ovf := #ovf);
	            "PDH_J_DTL"(v := #hbTs, zone := TRUE, buf := #pl, pos := #pos, ovf := #ovf);
	            "PDH_J_Raw"(s := ',"count":', buf := #pl, pos := #pos, ovf := #ovf);
	            "PDH_J_UDInt"(v := #heartbeatCount + 1, buf := #pl, pos := #pos, ovf := #ovf);
	            "PDH_J_Raw"(s := '}', buf := #pl, pos := #pos, ovf := #ovf);
	            #pubTopic := "PDH_Daten_Konfig".heartbeatTopic;
	            #pubRetain := FALSE;   // fest: ein alter Heartbeat darf nicht auf dem Broker liegen bleiben
	            // --- Ende Heartbeat ---
	    END_CASE;
	    IF NOT #ovf THEN
	        #pubLen := DINT_TO_UDINT(#pos);
	        #sendKind := #buildKind;
	        #pubReq := TRUE;   // steigende Flanke an publish im nächsten Aufruf
	        #state := 4;
	    ELSE
	        // Teil oder Heartbeat passt nicht: diesen Trigger verwerfen
	        #evStatus := 16#8008;
	        #evText := 'Nachricht zu lang';
	        IF #buildKind = 3 THEN
	            #hbDue := FALSE;
	        END_IF;
	        #busy := FALSE;
	        #state := 3;
	    END_IF;
	END_IF;

	// ---------------------------------------------------------------- Fehler: Bibliothek aus, 5 s warten, neu verbinden
	IF #failCode <> 16#0000 THEN
	    #failed := TRUE;
	    #lastErr := #failCode;
	    #lastText := #failText;
	    #connected := FALSE;
	    #busy := FALSE;
	    #trigPending := FALSE;
	    #hbDue := FALSE;
	    #pubReq := FALSE;
	    #libEnable := FALSE;
	    #state := 6;
	END_IF;

	// ---------------------------------------------------------------- Ausgänge
	IF #evStatus <> 16#0000 THEN
	    #error := TRUE;
	    #status := #evStatus;
	    #statusText := #evText;
	ELSIF #failed THEN
	    #error := TRUE;
	    #status := #lastErr;
	    #statusText := #lastText;
	ELSE
	    CASE #state OF
	        1:
	            IF #libStatus = 16#7003 THEN
	                #status := 16#7002;
	                #statusText := 'warte auf Broker';
	            ELSE
	                #status := 16#7001;
	                #statusText := 'verbinde';
	            END_IF;
	        3:
	            #status := 16#7003;
	            #statusText := 'bereit';
	        4:
	            IF #busy THEN
	                #status := 16#7004;
	                #statusText := 'sende';
	            ELSE
	                #status := 16#7003;
	                #statusText := 'bereit';
	            END_IF;
	        6:
	            IF #enable THEN
	                #status := 16#7001;
	                #statusText := 'verbinde';
	            ELSE
	                #status := 16#7000;
	                #statusText := 'aus';
	            END_IF;
	        ELSE
	            #status := 16#7000;
	            #statusText := 'aus';
	    END_CASE;
	END_IF;
END_FUNCTION_BLOCK

